// TIA Portal V20 export
Screen "150RobotCollision"  1276x673
  ScreenItem "Rectangle_4" at 160,488 size 164x112  Type=HmiRectangle
  ScreenItem "Rectangle_3" at 918,113 size 164x112  Type=HmiRectangle
  ScreenItem "矩形_6" at -3,69 size 1274x597  Type=HmiRectangle
  ScreenItem "Graphic view_13" at 324,99 size 634x531  Type=HmiGraphicView
  ScreenItem "Title_ScreenOverview_X390_Y2" at 438,5 size 551x57  Type=HmiTextBox
  ScreenItem "Line_Header_X0_Y64" at 0,64 size 1274x1  Type=HmiLine
  ScreenItem "permanentareaborderrectangle" at 0,0 size 0x0  Type=HmiRectangle
  ScreenItem "Button_Back" at 2,2 size 90x60  Type=HmiButton
  ScreenItem "Text_3" at 746,95 size 84x39  Type=HmiText
  ScreenItem "Text_4" at 734,600 size 84x39  Type=HmiText
  ScreenItem "Text_5" at 450,616 size 84x39  Type=HmiText
  ScreenItem "Text_6" at 461,80 size 84x39  Type=HmiText
  ScreenItem "Text_18" at 603,471 size 84x73  Type=HmiText
  ScreenItem "Graphic view_6" at 746,-206 size 60x30  Type=HmiGraphicView
  ScreenItem "Graphic view_7" at 746,-594 size 60x30  Type=HmiGraphicView
  ScreenItem "Graphic view_8" at 746,-982 size 60x30  Type=HmiGraphicView
  ScreenItem "Text_2" at 597,578 size 84x73  Type=HmiText
  ScreenItem "Rectangle_2" at 176,98 size 164x112  Type=HmiRectangle
  ScreenItem "Text_19" at 168,93 size 174x35  Type=HmiText
  ScreenItem "Text_20" at 199,119 size 123x35  Type=HmiText
  ScreenItem "Text_21" at 213,147 size 88x35  Type=HmiText
  ScreenItem "Text_22" at 205,175 size 136x35  Type=HmiText
  ScreenItem "矩形_8" at 189,182 size 17x17  Type=HmiRectangle
  ScreenItem "矩形_9" at 189,155 size 17x17  Type=HmiRectangle
  ScreenItem "矩形_10" at 189,128 size 17x17  Type=HmiRectangle
  ScreenItem "Graphic view_2" at 0,40 size 122x30  Type=HmiGraphicView
  ScreenItem "Graphic view_4" at 0,0 size 122x30  Type=HmiGraphicView
  ScreenItem "Text_1" at 603,75 size 84x73  Type=HmiText
  ScreenItem "Graphic view_1" at 0,40 size 122x30  Type=HmiGraphicView
  ScreenItem "Graphic view_3" at 0,0 size 122x30  Type=HmiGraphicView
  ScreenItem "Text_8" at 597,182 size 84x73  Type=HmiText
  ScreenItem "Text_7" at 947,190 size 136x35  Type=HmiText
  ScreenItem "矩形_11" at 931,197 size 17x17  Type=HmiRectangle
  ScreenItem "矩形_12" at 931,170 size 17x17  Type=HmiRectangle
  ScreenItem "Text_9" at 955,162 size 88x35  Type=HmiText
  ScreenItem "Text_23" at 941,134 size 123x35  Type=HmiText
  ScreenItem "矩形_13" at 931,143 size 17x17  Type=HmiRectangle
  ScreenItem "Text_24" at 910,108 size 174x35  Type=HmiText
  ScreenItem "Rectangle_1" at 918,457 size 164x112  Type=HmiRectangle
  ScreenItem "Text_10" at 947,534 size 136x35  Type=HmiText
  ScreenItem "矩形_1" at 931,541 size 17x17  Type=HmiRectangle
  ScreenItem "矩形_2" at 931,514 size 17x17  Type=HmiRectangle
  ScreenItem "Text_11" at 955,506 size 88x35  Type=HmiText
  ScreenItem "Text_12" at 941,478 size 123x35  Type=HmiText
  ScreenItem "矩形_3" at 931,487 size 17x17  Type=HmiRectangle
  ScreenItem "Text_13" at 910,452 size 174x35  Type=HmiText
  ScreenItem "Text_14" at 183,509 size 123x35  Type=HmiText
  ScreenItem "矩形_4" at 173,518 size 17x17  Type=HmiRectangle
  ScreenItem "Text_15" at 189,565 size 136x35  Type=HmiText
  ScreenItem "矩形_5" at 173,572 size 17x17  Type=HmiRectangle
  ScreenItem "矩形_7" at 173,545 size 17x17  Type=HmiRectangle
  ScreenItem "Text_16" at 197,537 size 88x35  Type=HmiText
  ScreenItem "Text_17" at 152,483 size 174x35  Type=HmiText
